Universal Robots URScript: TgtProg.script

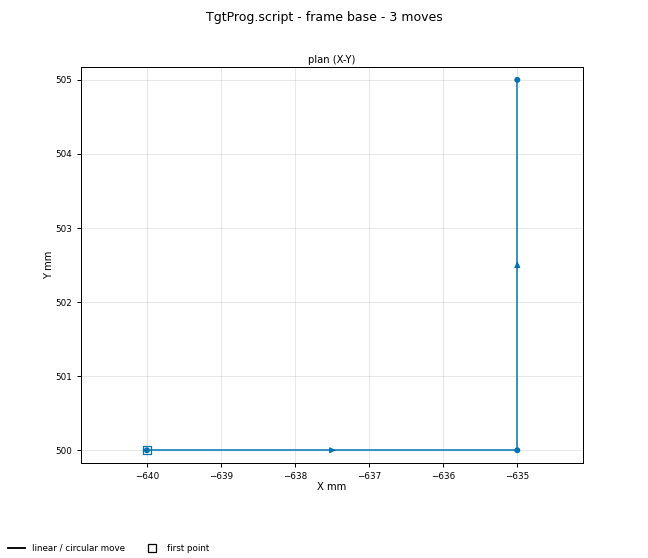
[picture p0: tool path of TgtProg.script in frame base, 3 of 3 moves have a stored position in this frame; points joined in program order, loops and branches not executed]
def TgtProg():
  # Global parameters:
  global speed_ms    = 0.250
  global speed_rads  = 0.750
  global accel_mss   = 1.200
  global accel_radss = 1.200
  global blend_radius_m = 0.001
  global ref_frame = p[0,0,0,0,0,0]

  #
  # TO REMOVE HEADER:
  # Go to "Program" -> "Post-Processor Editor"
  # Select "Universal Robots"
  # Set "INCLUDE_HEADER" to "False"
  #
  #--------------------------
  # Add any default subprograms here
  # For example, to drive a gripper as a program call:
  # def Gripper_Open():
  #   ...
  # end
  #
  # Example to drive a spray gun:
  def SprayOn(value):
    # use the value as an output:
    DO_SPRAY = 5
    if value == 0:
      set_standard_digital_out(DO_SPRAY, False)
    else:
      set_standard_digital_out(DO_SPRAY, True)
    end
  end

  # Example to drive an extruder:
  def Extruder(value):
    # use the value as an output:
    if value < 0:
      # stop extruder
    else:
      # start extruder
    end
  end

  # Example to move an external axis
  def MoveAxis(value):
    # use the value as an output:
    DO_AXIS_1 = 1
    DI_AXIS_1 = 1
    if value <= 0:
      set_standard_digital_out(DO_AXIS_1, False)

      # Wait for digital input to change state
      #while (get_standard_digital_in(DI_AXIS_1) != False):
      #  sync()
      #end
    else:
      set_standard_digital_out(DO_AXIS_1, True)

      # Wait for digital input to change state
      #while (get_standard_digital_in(DI_AXIS_1) != True):
      #  sync()
      #end
    end
  end
  #--------------------------


  # Main program:
  # Program generated by RoboDK v6.0.7 for UR10 on XX/XX/XXXX 18:00:00
  # Using nominal kinematics.
  blend_radius_m = 0.050
  movel(pose_trans(ref_frame,p[-0.640000, 0.500000, 0.370000, 0.731956, 2.185937, -0.570291]),accel_mss,speed_ms,t=0,r=0)
  movel(pose_trans(ref_frame,p[-0.635000, 0.500000, 0.370000, 0.731956, 2.185937, -0.570291]),accel_mss,speed_ms,t=0,r=0.050)
  movel(pose_trans(ref_frame,p[-0.635000, 0.505000, 0.370000, 0.731956, 2.185937, -0.570291]),accel_mss,speed_ms,t=0,r=0.050)
  # End of main program
end

TgtProg()
